TYPE "ST_LineRecord"
VERSION : 0.1
   STRUCT
      "WriteKey" : String[160];
      "Revision" : UDInt;
      "ValueText" : String[80];
   END_STRUCT;
END_TYPE
